Fanuc KAREL source: KT00854.KL

PROGRAM KT00854
%NOLOCKGROUP
VAR
  S1: STRING[80]
  S2: STRING[80]
  OUT: INTEGER
BEGIN
  S1 = 'A'
  S2 = 'B'
  S1 = 'A'
  S2 = 'B'
  OUT = TAN(S1)
END KT00854
